Universal Robots URScript: T012_mistralai_Devstral-Small-2-24B-Instruct-2512_baseline_rep1_retry2.urscript

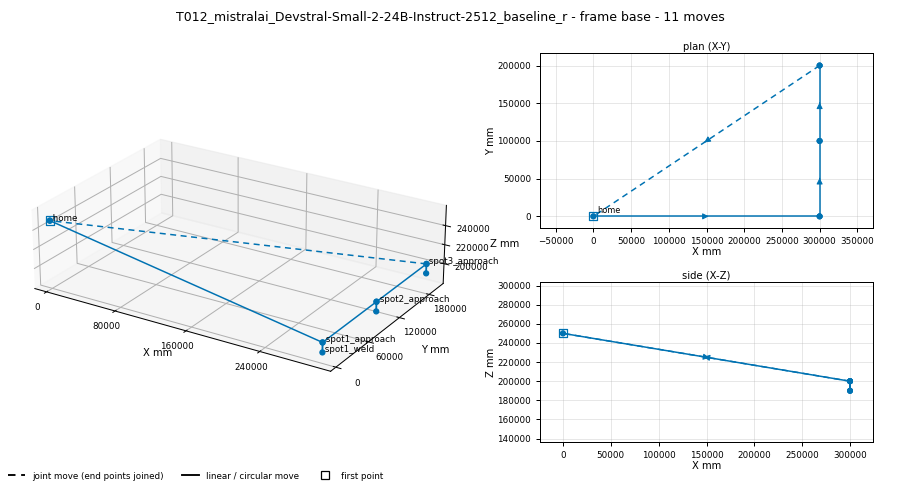
[picture p0: tool path of T012_mistralai_Devstral-Small-2-24B-Instruct-2512_baseline_rep1_retry2.urscript in frame base, 11 of 11 moves have a stored position in this frame; points joined in program order, loops and branches not executed]
def spot_welding():
    # Define tool and base frames
    tool0 = p[0, 0, 0, 0, 0, 0]
    base = p[0, 0, 0, 0, 0, 0]

    # Define spot positions (example coordinates)
    spot1_approach = p[300, 0, 200, 0, 0, 0]
    spot1_weld = p[300, 0, 190, 0, 0, 0]
    spot2_approach = p[300, 100, 200, 0, 0, 0]
    spot2_weld = p[300, 100, 190, 0, 0, 0]
    spot3_approach = p[300, 200, 200, 0, 0, 0]
    spot3_weld = p[300, 200, 190, 0, 0, 0]

    # Home position
    home = p[0, 0, 250, 0, 0, 0]

    # Set payload
    set_payload(2.5, p[0, 0, 0.1])

    # Set speed limits
    set_max_speed_l(250.0)
    set_max_speed_j(200.0)

    # Move to home position
    movej(home, a=1.4, v=200.0, t=0, r=0)

    # Spot 1
    movel(spot1_approach, a=1.4, v=200.0, t=0, r=0)
    movel(spot1_weld, a=1.4, v=80.0, t=0, r=0)
    # Simulate weld activation (replace with actual weld command)
    sleep(2.0)
    movel(spot1_approach, a=1.4, v=150.0, t=0, r=0)

    # Spot 2
    movel(spot2_approach, a=1.4, v=200.0, t=0, r=0)
    movel(spot2_weld, a=1.4, v=80.0, t=0, r=0)
    # Simulate weld activation
    sleep(2.0)
    movel(spot2_approach, a=1.4, v=150.0, t=0, r=0)

    # Spot 3
    movel(spot3_approach, a=1.4, v=200.0, t=0, r=0)
    movel(spot3_weld, a=1.4, v=80.0, t=0, r=0)
    # Simulate weld activation
    sleep(2.0)
    movel(spot3_approach, a=1.4, v=150.0, t=0, r=0)

    # Return to home
    movej(home, a=1.4, v=200.0, t=0, r=0)

spot_welding()
